Universal Robots URScript: T004_qwen2.5-coder_32b-instruct-q4_0_baseline_rep1.urscript

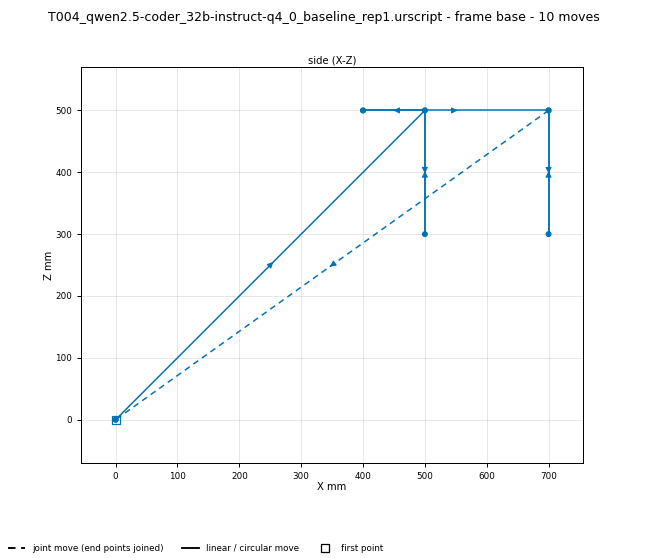
[picture p0: tool path of T004_qwen2.5-coder_32b-instruct-q4_0_baseline_rep1.urscript in frame base, 10 of 10 moves have a stored position in this frame; points joined in program order, loops and branches not executed]
# Multi-waypoint SSM pick-place with obstacle avoidance

# Home position
movej(p[0.0, -1.5708, 0.0, -1.5708, 0.0, 0.0], a=1.2, v=1.0, fine=TRUE)

# Move to WP1 - Above pick station
movel(p[0.5, -1.5708, 0.5, -1.5708, 0.0, 0.0], a=1.2, v=0.2)

# Move to WP2 - Descend to pick
movel(p[0.5, -1.5708, 0.3, -1.5708, 0.0, 0.0], a=1.2, v=0.1)

# Move to WP3 - Lift above pick
movel(p[0.5, -1.5708, 0.5, -1.5708, 0.0, 0.0], a=1.2, v=0.2)

# Move to WP4 - Obstacle avoidance waypoint (offset in -X)
movel(p[0.4, -1.5708, 0.5, -1.5708, 0.0, 0.0], a=1.2, v=0.2)

# Move to WP5 - Navigate around obstacle
movel(p[0.4, -1.5708, 0.5, -1.5708, 0.0, 0.5], a=1.2, v=0.2)

# Move to WP6 - Above place station
movel(p[0.7, -1.5708, 0.5, -1.5708, 0.0, 0.5], a=1.2, v=0.2)

# Move to WP7 - Descend to place
movel(p[0.7, -1.5708, 0.3, -1.5708, 0.0, 0.5], a=1.2, v=0.1)

# Move to WP8 - Lift above place
movel(p[0.7, -1.5708, 0.5, -1.5708, 0.0, 0.5], a=1.2, v=0.2)

# Return to Home position
movej(p[0.0, -1.5708, 0.0, -1.5708, 0.0, 0.0], a=1.2, v=1.0, fine=TRUE)
